{region 'Documentation'}
(*!
<summary>Checks reset reservation accounting on an exactly sized local Event Buffer.</summary>
<description>
Local counters represent two independent reservation callers, not child FB instances.
The budget is four Suite plus three Test Case entries and one shared Reset headroom.
Storage includes the FIFO spare position. These API tests do not prove owner admission.
Owner budget calculation and child dispatch are checked by separate integration scenarios.
The real subject binds only local storage; expected findings remain in that storage.
Checking Assertions retain the outer selftest publisher. Each run reinitializes the subject.
</description>
*)
{endregion}
FUNCTION_BLOCK Test_ResetReservationAccounting EXTENDS TestCaseBase
VAR
    FSubject : EventBuffer;
    FEvents : ARRAY[1..BufferLength] OF ST_Event;
    FFifo : ST_FifoStatus;
    FBufferStatus : ST_EventBufferStatus;
    FPerformed : BOOL;
    FChecked : BOOL;
    FSuiteReserved : UINT;
    FChildReserved : UINT;
    FInitialFifo : ST_FifoStatus;
    FBinding : AssertTrue;
    FBindingMatches : BOOL;
    FSuiteContribution : AssertTrue;
    FSuiteContributionMatches : BOOL;
    FCombinedContributions : AssertTrue;
    FCombinedContributionsMatches : BOOL;
    FRejectedReservation : AssertTrue;
    FRejectedReservationMatches : BOOL;
    FChildRelease : AssertTrue;
    FChildReleaseMatches : BOOL;
    FBalancedRelease : AssertTrue;
    FBalancedReleaseMatches : BOOL;
    FRepeatedRelease : AssertTrue;
    FRepeatedReleaseMatches : BOOL;
    FReadableDataUnchanged : AssertTrue;
    FReadableDataUnchangedMatches : BOOL;
END_VAR
VAR CONSTANT
    SuiteBudget : UINT := GVL_Constants.TestSuiteResetEventCount;
    ChildBudget : UINT := GVL_Constants.TestCaseResetEventCount;
    Headroom : UINT := Param_EventBuffer.EventBufferResetHeadroom;
    BufferLength : UINT := SuiteBudget + ChildBudget + Headroom + 1;
END_VAR

SUPER^();

{region 'Documentation'}
(*!
<summary>Contributes each checking Assertion once.</summary>
*)
{endregion}
METHOD PROTECTED AggregateResults
VAR_INPUT
    Aggregator : I_ResultAggregator; //! Borrowed result sink owned by the outer Test Case; add this test's checking Assertions without resetting or retaining the sink.
END_VAR
Aggregator.AddProvider(Provider := FBinding);
Aggregator.AddProvider(Provider := FSuiteContribution);
Aggregator.AddProvider(Provider := FCombinedContributions);
Aggregator.AddProvider(Provider := FRejectedReservation);
Aggregator.AddProvider(Provider := FChildRelease);
Aggregator.AddProvider(Provider := FBalancedRelease);
Aggregator.AddProvider(Provider := FRepeatedRelease);
Aggregator.AddProvider(Provider := FReadableDataUnchanged);
END_METHOD

{region 'Documentation'}
(*!
<summary>Requires all checking Assertions to be initialized.</summary>
*)
{endregion}
METHOD PROTECTED CheckInitialization : BOOL //! TRUE when the inherited initialization check and this concrete fixture check both accept the setup.
CheckInitialization := FALSE;
IF NOT SUPER^.CheckInitialization() THEN
    RETURN;
END_IF;

CheckInitialization := FBinding.IsInitialized
    AND FSuiteContribution.IsInitialized
    AND FCombinedContributions.IsInitialized
    AND FRejectedReservation.IsInitialized
    AND FChildRelease.IsInitialized
    AND FBalancedRelease.IsInitialized
    AND FRepeatedRelease.IsInitialized
    AND FReadableDataUnchanged.IsInitialized;
END_METHOD

{region 'Documentation'}
(*!
<summary>Initializes the checking Assertions for one test state.</summary>
*)
{endregion}
METHOD PROTECTED Configure
FPreparationStateCount := 0;
FTestStateCount := 1;
FBinding.Initialize(Parent := THIS^,
    AssertionName := 'Binding');
FSuiteContribution.Initialize(Parent := THIS^,
    AssertionName := 'SuiteContribution');
FCombinedContributions.Initialize(Parent := THIS^,
    AssertionName := 'CombinedContributions');
FRejectedReservation.Initialize(Parent := THIS^,
    AssertionName := 'RejectedReservation');
FChildRelease.Initialize(Parent := THIS^,
    AssertionName := 'ChildRelease');
FBalancedRelease.Initialize(Parent := THIS^,
    AssertionName := 'BalancedRelease');
FRepeatedRelease.Initialize(Parent := THIS^,
    AssertionName := 'RepeatedRelease');
FReadableDataUnchanged.Initialize(Parent := THIS^,
    AssertionName := 'ReadableDataUnchanged');
END_METHOD

{region 'Documentation'}
(*!
<summary>Checks local contributions and buffer-wide accounting at exact capacity.</summary>
*)
{endregion}
METHOD PRIVATE ExerciseBuffer
VAR
    Initialized : BOOL;
END_VAR
FSuiteReserved := 0;
FChildReserved := 0;
Initialized := FSubject.Initialize(Buffer := FEvents,
    FifoControl := FFifo,
    Status := FBufferStatus);
FBindingMatches := Initialized
    AND (FSubject.Capacity = BufferLength - 1)
    AND (FSubject.FreeEntryCount = BufferLength - 1)
    AND (FSubject.ReservedEntryCount = 0);
IF NOT Initialized THEN
    RETURN;
END_IF;

FInitialFifo := FFifo;
ReserveBudgets();
RejectAdditionalReservation();
ReleaseBudgets();

FReadableDataUnchangedMatches := (FFifo.IndexIn = FInitialFifo.IndexIn)
    AND (FFifo.IndexOut = FInitialFifo.IndexOut)
    AND (FFifo.ElementCount = 0) AND FFifo.BufferEmpty
    AND (FSubject.FreeEntryCount = BufferLength - 1)
    AND (FBufferStatus.SequenceId = 0)
    AND (FBufferStatus.DeletedSequenceId = 0)
    AND (FBufferStatus.LostEventCount = 0);
END_METHOD

{region 'Documentation'}
(*!
<summary>Completes abort without asynchronous work.</summary>
*)
{endregion}
METHOD PROTECTED ProcessAbort
VAR_INPUT
    Enable : BOOL; //! Phase permission supplied by the owning Test Case; FALSE does not authorize progression, while observation may continue.
END_VAR
IF Enable THEN
    CompleteAbort();
END_IF;
END_METHOD

{region 'Documentation'}
(*!
<summary>Evaluates captured observations after the scenario has finished.</summary>
*)
{endregion}
METHOD PROTECTED ProcessAssertions
VAR_INPUT
    Enable : BOOL; //! Phase permission supplied by the owning Test Case; FALSE does not authorize progression, while observation may continue.
END_VAR
VAR
    Evaluate : BOOL;
END_VAR
Evaluate := Enable AND FPerformed;
FBinding(Enable := Evaluate,
    State := State,
    IN := FBindingMatches);
FSuiteContribution(Enable := Evaluate,
    State := State,
    IN := FSuiteContributionMatches);
FCombinedContributions(Enable := Evaluate,
    State := State,
    IN := FCombinedContributionsMatches);
FRejectedReservation(Enable := Evaluate,
    State := State,
    IN := FRejectedReservationMatches);
FChildRelease(Enable := Evaluate,
    State := State,
    IN := FChildReleaseMatches);
FBalancedRelease(Enable := Evaluate,
    State := State,
    IN := FBalancedReleaseMatches);
FRepeatedRelease(Enable := Evaluate,
    State := State,
    IN := FRepeatedReleaseMatches);
FReadableDataUnchanged(Enable := Evaluate,
    State := State,
    IN := FReadableDataUnchangedMatches);
IF Evaluate THEN
    FChecked := TRUE;
END_IF;
END_METHOD

{region 'Documentation'}
(*!
<summary>No Preparation phase is needed.</summary>
*)
{endregion}
METHOD PROTECTED ProcessPreparations
VAR_INPUT
    // SA0033: Required override without Preparation work.
    {attribute 'analysis' := '-33'}
    Enable : BOOL; //! Phase permission supplied by the owning Test Case; FALSE does not authorize progression, while observation may continue.
END_VAR
END_METHOD

{region 'Documentation'}
(*!
<summary>Resets observations and schedules a fresh subject initialization.</summary>
*)
{endregion}
METHOD PROTECTED ProcessReset
FPerformed := FALSE;
FChecked := FALSE;
FBinding.Reset();
FBindingMatches := FALSE;
FSuiteContribution.Reset();
FSuiteContributionMatches := FALSE;
FCombinedContributions.Reset();
FCombinedContributionsMatches := FALSE;
FRejectedReservation.Reset();
FRejectedReservationMatches := FALSE;
FChildRelease.Reset();
FChildReleaseMatches := FALSE;
FBalancedRelease.Reset();
FBalancedReleaseMatches := FALSE;
FRepeatedRelease.Reset();
FRepeatedReleaseMatches := FALSE;
FReadableDataUnchanged.Reset();
FReadableDataUnchangedMatches := FALSE;
CompleteReset();
END_METHOD

{region 'Documentation'}
(*!
<summary>Runs the bounded scenario once before Assertion evaluation.</summary>
*)
{endregion}
METHOD PROTECTED ProcessTests
VAR_INPUT
    Enable : BOOL; //! Phase permission supplied by the owning Test Case; FALSE does not authorize progression, while observation may continue.
END_VAR
IF NOT Enable THEN
    RETURN;
END_IF;
IF FChecked THEN
    CompleteTests();
    RETURN;
END_IF;

IF NOT FPerformed THEN
    ExerciseBuffer();
    FPerformed := TRUE;
END_IF;
END_METHOD

{region 'Documentation'}
(*!
<summary>Verifies rejection leaves both contributions and the aggregate unchanged.</summary>
*)
{endregion}
METHOD PRIVATE RejectAdditionalReservation
VAR
    Accepted : BOOL;
END_VAR
Accepted := FSubject.ReserveSpace(EntryCount := 1,
    HeadroomEntryCount := Headroom,
    OwnerReservedEntryCount := FChildReserved);
FRejectedReservationMatches := NOT Accepted
    AND (FSuiteReserved = SuiteBudget) AND (FChildReserved = ChildBudget)
    AND (FSubject.ReservedEntryCount = SuiteBudget + ChildBudget);
END_METHOD

{region 'Documentation'}
(*!
<summary>Releases each contribution independently and repeats an empty release.</summary>
*)
{endregion}
METHOD PRIVATE ReleaseBudgets
VAR
    Released : BOOL;
END_VAR
Released := FSubject.FreeReservedSpace(EntryCount := FChildReserved,
    OwnerReservedEntryCount := FChildReserved);
FChildReleaseMatches := Released
    AND (FChildReserved = 0) AND (FSuiteReserved = SuiteBudget)
    AND (FSubject.ReservedEntryCount = SuiteBudget);

Released := FSubject.FreeReservedSpace(EntryCount := FSuiteReserved,
    OwnerReservedEntryCount := FSuiteReserved);
FBalancedReleaseMatches := Released
    AND (FSuiteReserved = 0) AND (FChildReserved = 0)
    AND (FSubject.ReservedEntryCount = 0);

Released := FSubject.FreeReservedSpace(EntryCount := FChildReserved,
    OwnerReservedEntryCount := FChildReserved);
FRepeatedReleaseMatches := Released
    AND (FChildReserved = 0) AND (FSuiteReserved = 0)
    AND (FSubject.ReservedEntryCount = 0);
END_METHOD

{region 'Documentation'}
(*!
<summary>Reserves two independent contributions with shared headroom.</summary>
*)
{endregion}
METHOD PRIVATE ReserveBudgets
VAR
    Accepted : BOOL;
END_VAR
Accepted := FSubject.ReserveSpace(EntryCount := SuiteBudget,
    HeadroomEntryCount := Headroom,
    OwnerReservedEntryCount := FSuiteReserved);
FSuiteContributionMatches := Accepted
    AND (FSuiteReserved = SuiteBudget) AND (FChildReserved = 0)
    AND (FSubject.ReservedEntryCount = SuiteBudget);

Accepted := FSubject.ReserveSpace(EntryCount := ChildBudget,
    HeadroomEntryCount := Headroom,
    OwnerReservedEntryCount := FChildReserved);
FCombinedContributionsMatches := Accepted
    AND (FSuiteReserved = SuiteBudget) AND (FChildReserved = ChildBudget)
    AND (FSubject.ReservedEntryCount = SuiteBudget + ChildBudget)
    AND (FSubject.FreeEntryCount = FSubject.ReservedEntryCount + Headroom);
END_METHOD

END_FUNCTION_BLOCK

(* stored: Version 1.1.0.1
   POU Test_ResetReservationAccounting: Id {feb0c693-aede-4cf9-9e73-372f2b368709}, SpecialFunc None
   Folder Internal: Id {cdbfd946-74ca-45a3-99c7-a33d730df0b5}
   Method AggregateResults: Id {64e3137c-ac17-4c09-aa90-a534c7f5eef6}
   Method CheckInitialization: Id {a8c245b8-fce2-425f-a98a-db4241316bdc}
   Method Configure: Id {b9432f04-62b4-42c5-80ba-247352bdd1e9}
   Method ExerciseBuffer: Id {69223444-ebd4-4e02-9d13-48fb01eec2d6}
   Method ProcessAbort: Id {7508e11d-b7a5-4586-a53e-2d2f283a108a}
   Method ProcessAssertions: Id {40f1b944-16e7-4ff2-8ccf-b96bc1caca82}
   Method ProcessPreparations: Id {7b7768a3-0ff8-43eb-a3c8-0bdb7069ec2c}
   Method ProcessReset: Id {e95cc33e-a08b-41d1-8278-1608a0f6e772}
   Method ProcessTests: Id {05dbcb3c-be18-4e85-91d1-fdfe479471ae}
   Method RejectAdditionalReservation: Id {e6c04d18-f8ad-45ff-9408-539c02382d05}
   Method ReleaseBudgets: Id {1e0fa68b-2de0-46a1-9394-aa498fd0de05}
   Method ReserveBudgets: Id {5f7afa97-a271-405b-8117-494f07a3e7b7} *)
